(*
SPDX-FileCopyrightText: © 2026 Oleksandr Tiutyk <trofimich@gmail.com>
SPDX-License-Identifier: MIT
License: https://opensource.org/license/mit
*)

(*!
<summary>Distinguishes execution-only, embedded and externally keyed bindings.</summary>
<description>Only embedded dependencies transfer ownership to the workflow.</description>
*)
{attribute 'qualified_only'}
{attribute 'strict'}
TYPE DEPENDENCY_BINDING_KIND :
(
	UNSPECIFIED,
	EMBEDDED,
	EXTERNAL_KEY
);
END_TYPE

(* stored: Version 1.1.0.1
   DUT DEPENDENCY_BINDING_KIND: Id {a70560a3-24d1-4d99-aea9-779db0febaf6} *)
